(* IEC 61131-3 sources: bevling_machine/framework/sources/01_Data, 8 files *)

(* ---- GVL_DeviceIds.st ---- *)
(* 模块说明：设备数组索引常量。D1..D8 对应索引 1..8，D6 保留；G1..G9 对应索引 9..17。

   全机所有设备数组共用这同一套 17 个索引，任何一处写错都会串到别人身上，所以先记住两条换算规则：
     D 编号 直接等于索引           D1..D8  ->  1..8
     G 编号 + 8 = 索引             G1..G9  ->  9..17

   ===== 17 个设备索引对照表 =====
   索引  代号  设备名称            类型       真实适配   绑定对象
   1     D1    送料皮带/输送轴     Axis       已接       songliao   点动/连续运行
   2     D2    切割走刀/回刀轴     Axis       已接       qiege      -
   3     D3    盘刀旋转电机        Axis       已接       pandao     按线性模式配置
   4     D4    定长平移轴          Axis       仿真       -          尚未接管
   5     D5    定长升降            Axis       仿真       -          0=升起避让，1=下降检测
   6     D6    定长光电            Sensor     已接       xDiMaterialLength 只读；TRUE=有料，遮挡即到位
   7     D7    机械手平移          Axis       仿真       -
   8     D8    平台旋转轴          Axis       已接       xuanzhuan  台达 ASDA-B3-E
   9     G1    下压气缸            Cylinder   已接       xDoG1ValveL/R  0=抬起，1=下压；左右双缸同动
   10    G2    侧挡升降（三缸）    Cylinder   已接       xDoG2Valve300/450/600 0=三缸全提，300/450/600=对应缸下降
   11    G3    推动气缸            Cylinder   已接       xDoG3Valve 0=放开，1=侧推
   12    G4    流利条升降          Cylinder   仿真       -          初始在提升端
   13    G5    喷油阀              Valve      仿真       xDoG5Spray 预留，待分配输出点
   14    G6    吹气阀              Valve      仿真       xDoG6Air   预留，待分配输出点
   15    G7    机械手升降          Cylinder   仿真       -          0=下降，1=提升
   16    G8    机械手夹爪          Cylinder   仿真       -          0=打开，1=夹紧
   17    G9    盘刀升降            Cylinder   已接       xDoG9Valve 0=提升，1=下降进刀

   报警码换算：整机报警 = 10000 + 索引。
     例：10001 = D1 皮带、10009 = G1 下压、10010 = G2 侧挡、10017 = G9 下刀。
     注意 10001 不是「1 号报警」，而是设备 1；真正的设备故障先看 udiErrorID 的千位。
   已在 FB_DeviceManager 中实现真实适配的编号：1、2、3、8（真实轴）、6（真实光电）与 9、10、11、17（真实气缸）。
   其余编号把 stReal.axRealDevice[i] 置 TRUE 会立即报 3002，不会被静默当仿真跑。 *)

VAR_GLOBAL CONSTANT
    D1_Belt : UINT := 1; (* D1 送料皮带电机，设备数组索引 1。 *)
    D2_CutFeed : UINT := 2; (* D2 切割走刀/回刀轴，设备数组索引 2。 *)
    D3_Spindle : UINT := 3; (* D3 盘刀旋转电机，设备数组索引 3。 *)
    D4_LengthMove : UINT := 4; (* D4 定长平移轴，设备数组索引 4。 *)
    D5_LengthLift : UINT := 5; (* D5 定长升降，0 升起避让，1 下降检测，索引 5。 *)
    D6_LengthSensor : UINT := 6; (* D6 定长光电（只读传感器），TRUE=有料，索引 6。 *)
    D7_GripperMove : UINT := 7; (* D7 机械手平移，索引 7；索引 6 为保留设备 D6。 *)
    D8_Rotate : UINT := 8; (* D8 平台旋转轴，设备数组索引 8。 *)
    G1_Press : UINT := 9; (* G1 下压气缸，0 抬起，1 下压，索引 9。 *)
    G2_SideStop : UINT := 10; (* G2 侧挡升降（三缸一组），目标 0=全提，300/450/600=对应缸下降，索引 10。 *)    (* G2 三个侧挡缸的料型号：同时作为设备 10 的命令目标值（lrTarget）和料型配方值（uiMaterialModel）。
       三者是同一套编号，不要再单独定义一套；界面上显示 300/450/600 就是这三个位号。 *)
    G2_Band300 : UINT := 300; (* G2 料型 300 对应的侧挡缸号。 *)
    G2_Band450 : UINT := 450; (* G2 料型 450 对应的侧挡缸号。 *)
    G2_Band600 : UINT := 600; (* G2 料型 600 对应的侧挡缸号。 *)
    G3_Push : UINT := 11; (* G3 推动气缸，0 放开，1 侧推，索引 11。 *)
    G4_RollerLift : UINT := 12; (* G4 流利条升降，0 下降，1 提升，索引 12。 *)
    G5_Spray : UINT := 13; (* G5 喷油阀，连续运行请求表示打开，索引 13。 *)
    G6_Air : UINT := 14; (* G6 吹气阀，切割开始打开、切割结束关闭，索引 14。 *)
    G7_GripperLift : UINT := 15; (* G7 机械手升降，0 下降，1 提升，索引 15。 *)
    G8_GripperClamp : UINT := 16; (* G8 机械手夹爪，0 打开，1 夹紧，索引 16。 *)
    G9_KnifeLift : UINT := 17; (* G9 盘刀升降，0 提升，1 下降，索引 17。 *)
END_VAR

(* ---- GVL_Interface.st ---- *)
(* 模块说明：监控与调试接口。stPanel 每周期由面板解码覆盖，不是上位机命令入口；手动请求保留待物理按钮映射。 *)
VAR_GLOBAL
    stPanel : ST_OperatorCommand; (* 本地面板解码结果，只读观察；每周期覆盖，操作请使用实体或仿真面板输入。 *)
    aManual : ARRAY[1..17] OF ST_ManualCommand; (* 各设备手动请求，索引 1..17；进入手动后先释放所有按钮再允许动作。 *)
    stStatus : ST_MachineStatus; (* 本模块对外发布的状态；字段含义见其数据类型。 *)
    aDeviceStatus : ARRAY[1..17] OF ST_DeviceStatus; (* 设备管理器汇总反馈，索引 1..17；供工序判断及在线监控。 *)
END_VAR

(* ---- GVL_IO.st ---- *)
(* 模块说明：逻辑 I/O 预留接口，尚未绑定物理地址。数字输出数组当前每周期清零；G2 当前料型仅用于观察。 *)
VAR_GLOBAL
    (* 当前均为普通逻辑变量，没有 AT %Q / %I 物理地址绑定。 *)
    xSafetyOK : BOOL; (* 安全许可接口或仿真许可，TRUE 允许；不等同于安全级急停回路。 *)
    stPanelInputs : ST_PanelInputs; (* 实体面板的模式旋钮、初始化、启动、停止、复位逻辑信号；急停走独立安全许可。 *)
    xMaterialAtLength : BOOL; (* 真实光电到位预留输入，当前未映射物理输入，仿真时不采用此值。 *)
    axDigitalInputs : ARRAY[0..31] OF BOOL; (* 预留数字输入位，索引 0..31；当前未映射到真实输入。 *)
    axDigitalOutputs : ARRAY[0..31] OF BOOL; (* 预留数字输出位，索引 0..31；当前由 FB_IOMap 每周期清 FALSE。 *)
    uiG2BandActive : UINT; (* G2 当前实际下降的料型带号 300/450/600；0 表示三缸全部提升，供诊断观察。 *)
END_VAR

(* ---- GVL_IO_Physical.st ---- *)
(* 模块说明：物理 I/O 符号层——传感器与电磁阀的唯一入口。
   本 GVL 刻意不带 AT %I* / AT %Q* 地址：通道由 InoProShop 的 I/O 映射页手工绑定，
   因此增减模块、调整 Local Bus 顺序都不会让符号与通道错位（地址由编译器重排，符号绑定不变）。

   极性约定（软件语义固定，与接线方式解耦）：
     DO  TRUE = 阀得电 = 设备动作（下压 / 伸出 / 下降）
     DI  TRUE = 该端到位
   若现场接线极性相反，只在本层取反，不改上层任何流程或互锁代码。

   当前分配建议（硬件工程师可调整，调整后同步改本注释即可）：
     DO  GL20_0032ETN  QB(I) bit0..bit4  -> G1左 / G1右 / G2-300 / G2-450 / G2-600
     DO  GL20_0032ETN  QB(I) bit5..bit6  -> G9 / 备用
     DO  指示灯另分配                    -> 绿灯 / 红灯
     DI  GL20_3200END  DI00..DI09        -> G1左(2) G2-300(2) G3(2) G9(2) G1右(2)
     DI  新增 4 点                       -> G2-450(2) G2-600(2)

   注意：G2 从单缸改成 300/450/600 三缸后，输出多占 2 点、输入多占 4 点。
   3200END 的 16 点 DI 原本已用 10 点，加 4 点后剩 2 点，仍然不够面板 8 点用，
   面板输入必须另加一块 DI 模块（这一点与改造前结论一致）。
   旧符号 xDoG2Valve / xDiG2Retract / xDiG2Extend 已停用，保留仅为避免已画好的
   映射页断开时报“符号不存在”，物理通道改绑到下方三个新阀与六个新限位符号。
*)
VAR_GLOBAL
    (* ===== 数字输出：GL20-0032ETN，单电控阀，高电平使能 ===== *)
    xDoG1ValveL : BOOL; (* G1 左压板阀：TRUE=下压，FALSE=抬起。建议 QB(I) bit0。 *)
    xDoG1ValveR : BOOL; (* G1 右压板阀：与左阀同命令同步动作。建议 QB(I) bit1。 *)
    xDoG2Valve300 : BOOL; (* G2 料型 300 侧挡阀：TRUE=该缸下降挡料，FALSE=提升。建议 QB(I) bit2。 *)
    xDoG2Valve450 : BOOL; (* G2 料型 450 侧挡阀：TRUE=该缸下降挡料，FALSE=提升。建议 QB(I) bit3。 *)
    xDoG2Valve600 : BOOL; (* G2 料型 600 侧挡阀：TRUE=该缸下降挡料，FALSE=提升。建议 QB(I) bit4。 *)
    xDoG3Valve : BOOL; (* G3 侧推阀：TRUE=侧推，FALSE=退回。建议 QB(I) bit5。 *)
    xDoG9Valve : BOOL; (* G9 盘刀升降阀：TRUE=下降进刀，FALSE=提升。建议 QB(I) bit6。 *)

    (* ===== 已停用：G2 原单缸阀。物理接线改绑 xDoG2Valve300/450/600，本符号保留不复用。 ===== *)
    xDoG2Valve : BOOL; (* 停用：G2 单缸阀旧符号，程序不再写入，保留仅为兼容已有映射页。 *)

    (* ===== 面板指示灯：两个纯输出，只有电平没有反馈 ===== *)
    xDoLampGreen : BOOL; (* 绿灯：手动/就绪常亮，自动循环运行中慢闪。 *)
    xDoLampRed : BOOL; (* 红灯：停机或故障时常亮。 *)

    (* ===== 数字输入：GL20-3200END，G1 双压板 4 点 + G3/G9 各 2 点 + G2 三缸 6 点 ===== *)
    (* G1 下压左压板 *)
    xDiG1LRetract : BOOL; (* 左缸抬起到位。建议 DI00。 *)
    xDiG1LExtend : BOOL; (* 左缸下压到位。建议 DI01。 *)

    (* G2 侧挡 300 缸 *)
    xDiG2_300Retract : BOOL; (* 300 缸提升到位。建议 DI02。 *)
    xDiG2_300Extend : BOOL; (* 300 缸下降到位。建议 DI03。 *)

    (* G3 侧推气缸 *)
    xDiG3Retract : BOOL; (* G3 退回到位。建议 DI04。 *)
    xDiG3Extend : BOOL; (* G3 伸出到位。建议 DI05。 *)

    (* G9 盘刀升降 *)
    xDiG9Retract : BOOL; (* G9 提升到位。建议 DI06。 *)
    xDiG9Extend : BOOL; (* G9 下降到位。建议 DI07。 *)

    (* G1 下压右压板：与左压板同属设备索引 9，两组传感器必须同时到位才算该端到位 *)
    xDiG1RRetract : BOOL; (* 右缸抬起到位。建议 DI08。 *)
    xDiG1RExtend : BOOL; (* 右缸下压到位。建议 DI09。 *)

    (* G2 侧挡 450 / 600 缸：新增 4 点，3200END 已无空位，需另加 DI 模块或换 32 点模块 *)
    xDiG2_450Retract : BOOL; (* 450 缸提升到位。 *)
    xDiG2_450Extend : BOOL; (* 450 缸下降到位。 *)
    xDiG2_600Retract : BOOL; (* 600 缸提升到位。 *)
    xDiG2_600Extend : BOOL; (* 600 缸下降到位。 *)

    (* ===== 已停用：G2 原单缸限位。改用上方三缸各自的六个限位符号。 ===== *)
    xDiG2Retract : BOOL; (* 停用：G2 单缸提升到位旧符号，程序不再读取。 *)
    xDiG2Extend : BOOL; (* 停用：G2 单缸下降到位旧符号，程序不再读取。 *)

    (* ===== 定长光电：D6，遮挡=有料。通道由映射页手工绑定，接哪个模块哪一位都行 ===== *)
    xDiMaterialLength : BOOL; (* 定长光电：TRUE=被遮挡=料已到位。建议接在还空着的 DI 上。 *)

    (* ===== 预留：喷油 / 吹气（本轮不接，占位避免后期改结构） ===== *)
    xDoG5Spray : BOOL; (* 喷油阀：TRUE=喷油。待分配。 *)
    xDoG6Air : BOOL; (* 吹气阀：TRUE=吹气。待分配。 *)

    (* ===== 测试控制面板输入：符号名固定，通道同样由映射页手工绑定 ===== *)
    (* 极性：除急停与停止外，均为常开触点，按下/到位为 TRUE。 *)
    xDiPanelAutoMode : BOOL; (* 自动/手动旋钮：TRUE=自动，FALSE=手动。 *)
    xDiPanelSafetyPermit : BOOL; (* 安全许可旋钮：TRUE=许可。 *)
    xDiEStop : BOOL; (* 急停自锁按钮，常开，按下=TRUE=不安全；断线读 FALSE 软件无法分辨，需外部安全回路。 *)
    xDiPanelRunStart : BOOL; (* 启动按钮，常开，按下=TRUE；上升沿把整机置为运行态。 *)
    xDiPanelRunStop : BOOL; (* 停止按钮，常闭：未按=TRUE，按下=FALSE；逻辑层取反后按上升沿处理。 *)
    xDiPanelStart : BOOL; (* start 按钮，常开，按下=TRUE；自动循环启动，须已初始化到 Ready。 *)
    xDiPanelInit : BOOL; (* 初始化按钮，常开，按下=TRUE。 *)
    xDiPanelReset : BOOL; (* 报警复位按钮，常开，按下=TRUE。 *)
END_VAR

(* ---- GVL_Modbus.st ---- *)
(* 模块说明：Modbus 收发缓冲区，索引从 0 开始，尚未绑定网络寄存器。实际地址和字序需另行配置。 *)
VAR_GLOBAL
    (* 仅预留收发缓冲区，尚未绑定工程中的 MODBUS_TCP 网络映射。 *)
    xEnable : BOOL; (* 启用 Modbus 缓冲区解析，默认 FALSE；不代表网络映射已经配置。 *)
    awRx : ARRAY[0..31] OF WORD; (* v2 接收字：0=版本2，1=序号，2=命令2启动/3停止；3/4 保留且必须为0，不接受模式写入。 *)
    awTx : ARRAY[0..127] OF WORD; (* 发布字缓冲区 0..127；包含确认、状态、报警、计数和位置，详见程序内索引注释。 *)
END_VAR

(* ---- GVL_Parameters.st ---- *)
(* 模块说明：仿真开关和待执行配方。参数生效时机见 ST_Recipe；关闭仿真当前报 3001，未接入真实设备。 *)
VAR_GLOBAL
    (* 以下默认值仅供软件仿真，不能直接作为已确认的生产参数。 *)
    xSimulation : BOOL := TRUE; (* TRUE 使用内部仿真；当前 FALSE 报未实现 3001，不会接管真实运动。 *)
    xContinuous : BOOL := FALSE; (* 本地工程配置的单循环/连续选择；上位机启停帧不修改此设置，默认单循环。 *)
    xAllowRemoteStartStop : BOOL := FALSE; (* 本地工程配置授权远程启停，默认 FALSE；不授予改模式、初始化或复位权限，也不映射给上位机写。 *)
    stRecipe : ST_Recipe; (* 待执行配方：初始化和自动启动时校验并取快照，运行中修改不会立即生效。 *)
    xUseRealPanel : BOOL := TRUE; (* TRUE 读物理面板按钮/旋钮；FALSE 读仿真面板。与 xSimulation 解耦，后者恒为 TRUE。 *)
END_VAR

(* ---- GVL_RealDevice.st ---- *)
(* 模块说明：真实设备接管设置的唯一入口。默认全部 FALSE，整机行为与改造前完全一致。 *)
VAR_GLOBAL
	stSettings : ST_RealDeviceSettings; (* 接管开关、验证参数、旁路开关集中在此，便于 HMI 与调试统一读写。 *)
END_VAR

(* ---- GVL_Simulation.st ---- *)
(* 模块说明：仿真调试入口。可模拟来料、动作卡住、设备故障和安全许可丢失。 *)
VAR_GLOBAL
    stSettings : ST_SimulationSettings; (* 软件仿真参数，含来料方式和异常注入。 *)
    stPanelInputs : ST_PanelInputs; (* 仿真旋钮/按钮输入；xAutoMode 选择模式，其余按钮按住/释放模拟物理信号。 *)
END_VAR
